Fanuc KAREL source: KA00225.KL

PROGRAM KA00225
%NOLOCKGROUP
VAR
  SRC: ARRAY[4] OF JOINTPOS
  DST: ARRAY[4] OF JOINTPOS
BEGIN
  DST = SRC
END KA00225
